Staubli VAL3: action.pjx

--- action.pjx ---
Parameters version=s8.10.3Cs9_BS2093 stackSize=5000 millimeterUnit=true
Program file=start.pgx
Program file=stop.pgx
Data file=action.dtx

--- action.dtx ---
public num nActResult
public num nActType
public num nActIO

--- start.pgx ---
program start()
begin
end

--- stop.pgx ---
program stop()
begin
end
